(* PLC project Storage_Main, Beckhoff Automation GmbH TwinCAT PLC Control 3.5.13.21 *)
(* stored: creationDateTime 2026-11-24T10:23:53.5609377, modificationDateTime 2026-11-24T10:23:53.5609377 *)

PROGRAM MAIN
// =====================================================================
// MAIN (Structured Text)
// Calls the ST actions and the SFC action ACT_Sequence in a fixed order.
// All variables of the storage system are declared here (HMI uses MAIN.xxx).
// =====================================================================
VAR
    // ---------------- INPUTS ----------------
    B1  AT %I* : BOOL;  // Nr. 5,  B1: reference switch horizontal axis (TRUE = at home)
    B2  AT %I* : BOOL;  // Nr. 6,  B2: light-barrier inside  (TRUE = free, FALSE = pallet)
    B3  AT %I* : BOOL;  // Nr. 7,  B3: light-barrier outside (TRUE = free, FALSE = pallet)
    B4  AT %I* : BOOL;  // Nr. 8,  B4: reference switch vertical axis, top (TRUE = at home)
    B5  AT %I* : BOOL;  // Nr. 11, B5: encoder horizontal axis impulse 1  (EL1202 Term 2 ch. 1)
    B6  AT %I* : BOOL;  // Nr. 12, B6: encoder horizontal axis impulse 2  (EL1202 Term 2 ch. 2)
    B7  AT %I* : BOOL;  // Nr. 13, B7: encoder vertical axis impulse 1    (EL1202 Term 3 ch. 1)
    B8  AT %I* : BOOL;  // Nr. 14, B8: encoder vertical axis impulse 2    (EL1202 Term 3 ch. 2)
    B9  AT %I* : BOOL;  // Nr. 15, B9: reference switch cantilever front (TRUE = arm out)
    B10 AT %I* : BOOL;  // Nr. 16, B10: reference switch cantilever back (TRUE = arm back)

    // ---------------- OUTPUTS ----------------
    M1_Forward AT %Q* : BOOL;  // Nr. 17, Q1 (M1): motor conveyor belt forward
    M1_Back    AT %Q* : BOOL;  // Nr. 18, Q2 (M1): motor conveyor belt backward (moves pallet towards crane)
    M2_Forward AT %Q* : BOOL;  // Nr. 19, Q3 (M2): motor horizontal towards rack
    M2_Back    AT %Q* : BOOL;  // Nr. 20, Q4 (M2): motor horizontal towards conveyor belt
    M3_Down    AT %Q* : BOOL;  // Nr. 21, Q5 (M3): motor vertical axis downward
    M3_Up      AT %Q* : BOOL;  // Nr. 22, Q6 (M3): motor vertical axis upward
    M4_Forward AT %Q* : BOOL;  // Nr. 23, Q7 (M4): motor cantilever forward (arm out)
    M4_Back    AT %Q* : BOOL;  // Nr. 24, Q8 (M4): motor cantilever backward (arm in)

    nTolerance   : DINT := 5;       // Deadband in counts (both axes)

    // ---------------- MANUAL COMMANDS (step S0 only) ----------------
    bJogXForward    : BOOL;         // X towards rack
    bJogXBack       : BOOL;         // X towards conveyor
    bJogYUp         : BOOL;         // Y up
    bJogYDown       : BOOL;         // Y down
    bJogArmOut      : BOOL;         // Arm out (stops at B9)
    bJogArmIn       : BOOL;         // Arm in (stops at B10)
    bJogBeltForward : BOOL;         // Belt moves pallet towards crane (M1_Back, stops when B3 sees a pallet)
    bJogBeltBack    : BOOL;         // Belt moves pallet away from crane (M1_Forward)

    // ---------------- TEACH ----------------
    nTeachSlot : INT := 0;          // 0 = delivery (conveyor), 1..3 = column (X) / row (Y)
    bTeachX    : BOOL;              // Save nPosX into xPosition[nTeachSlot]
    bTeachY    : BOOL;              // Save nPosY into yPosition[nTeachSlot]
    bGoX       : BOOL;              // Move X to xPosition[nTeachSlot]
    bGoY       : BOOL;              // Move Y to yPosition[nTeachSlot]
    nShowX     : DINT;              // Stored X value of nTeachSlot (for HMI)
    nShowY     : DINT;              // Stored Y value of nTeachSlot (for HMI)

    // ---------------- SAVE TAUGHT VALUES (Tc2_Utilities) ----------------
    fbWritePersistent : WritePersistentData;   // Writes all PERSISTENT variables to disk at once
    bSaveData         : BOOL;       // Request: save the persistent data now
    nSaveState        : INT;        // 0 = idle, 1 = start writing, 2 = writing
    bSaveError        : BOOL;       // TRUE if the last write failed
    nLiftOffsetOld    : DINT;       // Last saved nLiftOffset (detects a change from the HMI)
    nLowerOffsetOld   : DINT;       // Last saved nLowerOffset (detects a change from the HMI)

    // ---------------- AUTOMATIC ----------------
    bStartAuto     : BOOL;          // Start automatic mode (homes first)
    bStartHoming   : BOOL;          // Start homing (manual mode)
    bStop          : BOOL;          // Stop everything, back to manual
    bAuto          : BOOL;          // TRUE while automatic mode is active
    bResetSequence : BOOL;          // TRUE for one cycle: ACT_Sequence back to step S0 (STOP / homing timeout)
    SFCReset       : BOOL;          // SFC flag of ACT_Sequence (set from bResetSequence in MAIN)
    nSelColumn     : INT;           // Shelf column to fetch from, chosen by the operator (1..3)
    nSelRow        : INT;           // Shelf row to fetch from, chosen by the operator (1..3)
    bShelfSelected : BOOL;          // Set by the HMI when the operator has chosen a shelf
    bPositionFound : BOOL;          // GRAFCET: PositionFound - target position is loaded (step 71 / 79)
    bInPosition    : BOOL;          // GRAFCET: InPosition - both axes are in position (step 77 / 84)

    // ---------------- POSITIONING ----------------
    nTargetX     : DINT;            // Current X target (GRAFCET: PosX value)
    nTargetY     : DINT;            // Current Y target (GRAFCET: PosY value)
    bDriveX      : BOOL;            // Sequence requests X to move to nTargetX
    bDriveY      : BOOL;            // Sequence requests Y to move to nTargetY
    bPosXReached : BOOL;            // GRAFCET: PosX = TRUE - X has reached nTargetX
    bPosYReached : BOOL;            // GRAFCET: PosY = TRUE - Y has reached nTargetY

    // ---------------- LIMITS ----------------
    nMaxPosX     : DINT := 10000;   // Software end limit X towards rack - MEASURE THIS!
    nMaxPosY     : DINT := 10000;   // Software end limit Y downwards - MEASURE THIS!
    tonHoming    : TON;             // Homing timeout
    bHomingError : BOOL;            // TRUE if a reference switch was not found in time
    tonSettle    : TON;             // 0.5 s settle time at the reference switches

    // ---------------- ENCODER X (B5/B6) ----------------
    nStateX      : BYTE;            // Current state 0..3
    nPrevStateX  : BYTE;            // State in previous cycle
    nPosX        : DINT;            // X position in counts (0 = B1, increases towards rack)
    nErrorCountX : UDINT;           // Number of missed states X

    // ---------------- ENCODER Y (B7/B8) ----------------
    nStateY      : BYTE;            // Current state 0..3
    nPrevStateY  : BYTE;            // State in previous cycle
    nPosY        : DINT;            // Y position in counts (0 = B4 at the top, increases downwards)
    nErrorCountY : UDINT;           // Number of missed states Y

    bInit : BOOL := TRUE;           // First cycle flag (both encoders)

    // ---------------- SEQUENCE / STATUS ----------------
    nStep            : INT := 0;    // Active SFC step number (set by the step actions of ACT_Sequence)
    bHomed           : BOOL;        // TRUE when both axes are homed
    bYTaught         : BOOL;        // TRUE when all Y positions are taught
    bYNotTaught      : BOOL;        // Inverse of bYTaught (for HMI)
    bPalletAtB2      : BOOL;        // TRUE when B2 sees a pallet (HMI lamp)
    bPalletAtB3      : BOOL;        // TRUE when B3 sees a pallet (HMI lamp)
    bShowShelfSelect : BOOL;        // TRUE while the operator must choose a shelf (shows 3x3 on HMI)
    bHideShelfSelect : BOOL;        // Inverse of bShowShelfSelect (hides the 3x3 frame on HMI)
    bSlot0Sel        : BOOL;        // TRUE when teach slot 0 (delivery) is selected (lights the HMI button)
    bSlot1Sel        : BOOL;        // TRUE when teach slot 1 (column 1 / row 1) is selected
    bSlot2Sel        : BOOL;        // TRUE when teach slot 2 (column 2 / row 2) is selected
    bSlot3Sel        : BOOL;        // TRUE when teach slot 3 (column 3 / row 3) is selected
END_VAR

VAR PERSISTENT
    // ---------------- TAUGHT VALUES (kept after power off) ----------------
    // Index 0 = delivery position at the conveyor (GRAFCET: DeliveryPosX / DeliveryPosY)
    // X: [1] = column 1 (nearest conveyor) .. [3] = column 3
    // Y: [1] = row 1 (bottom) .. [3] = row 3 (top). Y counts from the top (B4 = 0) and increases downwards
    xPosition    : ARRAY[0..3] OF DINT := [139, 2995, 5330, 7680];
    yPosition    : ARRAY[0..3] OF DINT := [0, 0, 0, 0];      // MUST BE TAUGHT before automatic mode
    nLiftOffset  : DINT := 30;      // Counts to lift the pallet off the shelf (SFC step S74)
    nLowerOffset : DINT := 50;      // Counts to lower the pallet onto the conveyor (SFC step S86)
END_VAR

            // =====================================================================
// MAIN (Structured Text) - the order of the calls is important:
//   1. ACT_Encoder     (ST)  read the encoders -> nPosX / nPosY
//   2. ACT_Manual      (ST)  status, stop, commands, teach + save, timers,
//                            all motors off, jog in manual mode
//   3. ACT_Sequence    (SFC) homing and the automatic sequence (switches motors ON)
//   4. ACT_Positioning (ST)  drive X / Y to nTargetX / nTargetY
//   5. ACT_Safety      (ST)  end limits and interlocks (always last)
// =====================================================================

ACT_Encoder();
ACT_Manual();

SFCReset := bResetSequence;                 // SFC flag: TRUE = ACT_Sequence back to step S0
ACT_Sequence();                             // SFC: homing and automatic sequence
bResetSequence := FALSE;

// Commands are only accepted in manual mode (step S0). Clear them every cycle,
// so an old button press does not start something later by surprise.
bStartHoming := FALSE;
bStartAuto   := FALSE;
bGoX         := FALSE;
bGoY         := FALSE;

ACT_Positioning();
ACT_Safety();

          

ACTION ACT_Encoder:
                // =====================================================
// ACT_Encoder: count up/down based on the two encoder signals
// X: B5 (A) and B6 (B)    Y: B7 (A) and B8 (B)
// =====================================================
nStateX := 0;                                       // default: A=0, B=0
IF B5 AND NOT B6 THEN nStateX := 1; END_IF          // A=1, B=0
IF B5 AND B6 THEN nStateX := 2; END_IF              // A=1, B=1
IF NOT B5 AND B6 THEN nStateX := 3; END_IF          // A=0, B=1

nStateY := 0;                                       // default: A=0, B=0
IF B7 AND NOT B8 THEN nStateY := 1; END_IF          // A=1, B=0
IF B7 AND B8 THEN nStateY := 2; END_IF              // A=1, B=1
IF NOT B7 AND B8 THEN nStateY := 3; END_IF          // A=0, B=1

IF bInit THEN
    nPrevStateX := nStateX;
    nPrevStateY := nStateY;
    bInit := FALSE;
END_IF

CASE (nStateX + 4 - nPrevStateX) MOD 4 OF
    1: nPosX := nPosX + 1;                          // one step towards rack
    3: nPosX := nPosX - 1;                          // one step towards conveyor
    2: nErrorCountX := nErrorCountX + 1;            // state missed
END_CASE

CASE (nStateY + 4 - nPrevStateY) MOD 4 OF
    1: nPosY := nPosY + 1;                          // one step down
    3: nPosY := nPosY - 1;                          // one step up
    2: nErrorCountY := nErrorCountY + 1;            // state missed
END_CASE

nPrevStateX := nStateX;
nPrevStateY := nStateY;

              
END_ACTION

ACTION ACT_Manual:
                // =====================================================
// ACT_Manual: status, stop, commands, teach + save, timers, jog
// =====================================================

// ---------- 1. STATUS SIGNALS ----------
bPalletAtB2 := NOT B2;                              // light barrier is FALSE when a pallet is in front
bPalletAtB3 := NOT B3;

// Delivery height must be taught, and every shelf row must be low enough to lift nLiftOffset
bYTaught := yPosition[0] > 0 AND yPosition[1] > nLiftOffset AND yPosition[2] > nLiftOffset AND yPosition[3] > nLiftOffset;
bYNotTaught := NOT bYTaught;

bShowShelfSelect := (nStep = 71);
bHideShelfSelect := NOT bShowShelfSelect;
bSlot0Sel := (nTeachSlot = 0);
bSlot1Sel := (nTeachSlot = 1);
bSlot2Sel := (nTeachSlot = 2);
bSlot3Sel := (nTeachSlot = 3);

IF nTeachSlot >= 0 AND nTeachSlot <= 3 THEN
    nShowX := xPosition[nTeachSlot];
    nShowY := yPosition[nTeachSlot];
END_IF


// ---------- 2. STOP: always back to manual mode (step S0) ----------
IF bStop THEN
    bStop := FALSE;
    bStartHoming := FALSE;
    bStartAuto := FALSE;
    bGoX := FALSE;
    bGoY := FALSE;
    bShelfSelected := FALSE;
    bPositionFound := FALSE;
    bInPosition := FALSE;
    bAuto := FALSE;
    bResetSequence := TRUE;                         // ACT_Sequence -> S0 (SFCReset)
END_IF


// ---------- 3. COMMANDS (manual mode only) ----------
// The transitions after step S0 in ACT_Sequence react to the same commands in this cycle.
IF nStep = 0 THEN
    IF bStartHoming THEN
        bHomingError := FALSE;
        bAuto := FALSE;
        bHomed := FALSE;
    END_IF

    IF bStartAuto AND bYTaught THEN                 // Y positions must be taught first
        bHomingError := FALSE;
        bAuto := TRUE;
        bHomed := FALSE;                            // always home before automatic mode
    END_IF

    IF bGoX AND bHomed AND nTeachSlot >= 0 AND nTeachSlot <= 3 THEN
        nTargetX := xPosition[nTeachSlot];
        bPosXReached := FALSE;
    END_IF

    IF bGoY AND bHomed AND nTeachSlot >= 0 AND nTeachSlot <= 3 THEN
        nTargetY := yPosition[nTeachSlot];
        bPosYReached := FALSE;
    END_IF
END_IF


// ---------- 4. TEACH: save current position into the arrays (manual mode only) ----------
IF bTeachX THEN
    bTeachX := FALSE;
    IF nStep = 0 AND bHomed AND nTeachSlot >= 0 AND nTeachSlot <= 3 THEN
        xPosition[nTeachSlot] := nPosX;
        bSaveData := TRUE;                          // write to disk at once
    END_IF
END_IF

IF bTeachY THEN
    bTeachY := FALSE;
    IF nStep = 0 AND bHomed AND nTeachSlot >= 0 AND nTeachSlot <= 3 THEN
        yPosition[nTeachSlot] := nPosY;
        bSaveData := TRUE;                          // write to disk at once
    END_IF
END_IF

// Lift / lower offset changed on the HMI -> save as well
IF nLiftOffset <> nLiftOffsetOld OR nLowerOffset <> nLowerOffsetOld THEN
    nLiftOffsetOld := nLiftOffset;
    nLowerOffsetOld := nLowerOffset;
    bSaveData := TRUE;
END_IF


// ---------- 5. SAVE: write the PERSISTENT variables to disk (survives a power cut) ----------
// WritePersistentData starts on a rising edge of START. nSaveState makes sure that
// START is TRUE until the write has started, and FALSE again before the next write.
CASE nSaveState OF
    0:  // idle: wait for a save request
        IF bSaveData THEN
            bSaveData := FALSE;
            nSaveState := 1;
        END_IF

    1:  // START = TRUE: wait until the write has started (or failed at once)
        IF fbWritePersistent.BUSY OR fbWritePersistent.ERR THEN
            nSaveState := 2;
        END_IF

    2:  // START = FALSE: wait until the write is finished
        IF NOT fbWritePersistent.BUSY THEN
            nSaveState := 0;
        END_IF
END_CASE

fbWritePersistent(NETID := '', PORT := 851, START := (nSaveState = 1), TMOUT := T#5S, MODE := SPDM_2PASS);
bSaveError := fbWritePersistent.ERR;


// ---------- 6. TIMERS (called every cycle so they reset themselves) ----------
tonHoming(IN := (nStep = 10 OR nStep = 11), PT := T#20S);
tonSettle(IN := (nStep = 12), PT := T#500MS);

IF tonHoming.Q THEN
    bHomingError := TRUE;
    bAuto := FALSE;
    bResetSequence := TRUE;                         // ACT_Sequence -> S0, motors off
END_IF


// ---------- 7. MOTORS OFF + JOG ----------
// Default: all motors off. ACT_Sequence (called after this action) switches on what
// the active step needs. In manual mode (S0) the jog buttons are used.
M1_Forward := FALSE;
M1_Back    := FALSE;
M2_Forward := FALSE;
M2_Back    := FALSE;
M3_Down    := FALSE;
M3_Up      := FALSE;
M4_Forward := FALSE;
M4_Back    := FALSE;
bDriveX    := FALSE;
bDriveY    := FALSE;

IF nStep = 0 THEN
    M2_Forward := bJogXForward AND NOT bJogXBack;
    M2_Back    := bJogXBack AND NOT bJogXForward;
    M3_Down    := bJogYDown AND NOT bJogYUp;
    M3_Up      := bJogYUp AND NOT bJogYDown;
    M4_Forward := bJogArmOut AND NOT bJogArmIn;
    M4_Back    := bJogArmIn AND NOT bJogArmOut;
    M1_Back    := bJogBeltForward AND NOT bJogBeltBack AND B3;   // stops when B3 sees a pallet
    M1_Forward := bJogBeltBack AND NOT bJogBeltForward;
END_IF

              
END_ACTION

ACTION ACT_Positioning:
                // =====================================================
// ACT_Positioning: drive X and Y to their targets
// =====================================================
// An axis stops for good when it is within the tolerance (bPosXReached / bPosYReached),
// so it does not hunt back and forth if the motor coasts a little.
IF bDriveX AND NOT bPosXReached THEN
    IF nPosX < nTargetX - nTolerance THEN
        M2_Forward := TRUE;                         // towards rack
    END_IF
    IF nPosX > nTargetX + nTolerance THEN
        M2_Back := TRUE;                            // towards conveyor
    END_IF
    IF NOT M2_Forward AND NOT M2_Back THEN
        bPosXReached := TRUE;
    END_IF
END_IF

IF bDriveY AND NOT bPosYReached THEN
    IF nPosY < nTargetY - nTolerance THEN
        M3_Down := TRUE;                            // larger Y = further down
    END_IF
    IF nPosY > nTargetY + nTolerance THEN
        M3_Up := TRUE;                              // smaller Y = further up
    END_IF
    IF NOT M3_Down AND NOT M3_Up THEN
        bPosYReached := TRUE;
    END_IF
END_IF

              
END_ACTION

ACTION ACT_Safety:
                // =====================================================
// ACT_Safety: end limits and interlocks (always called last)
// =====================================================
// X: hardware end at the conveyor (B1)
IF B1 THEN
    M2_Back := FALSE;
END_IF

// X: software end towards the rack
IF bHomed AND nPosX >= nMaxPosX THEN
    M2_Forward := FALSE;
END_IF

// X may only move when the arm is back (B10)
IF NOT B10 THEN
    M2_Forward := FALSE;
    M2_Back    := FALSE;
END_IF

// Y: hardware end at the top (B4)
IF B4 THEN
    M3_Up := FALSE;
END_IF

// Y: software end at the bottom
IF bHomed AND nPosY >= nMaxPosY THEN
    M3_Down := FALSE;
END_IF

// Arm: end positions
IF B9 THEN
    M4_Forward := FALSE;
END_IF

IF B10 THEN
    M4_Back := FALSE;
END_IF

// Never both directions at the same time
IF M1_Forward AND M1_Back THEN
    M1_Forward := FALSE;
    M1_Back    := FALSE;
END_IF

IF M2_Forward AND M2_Back THEN
    M2_Forward := FALSE;
    M2_Back    := FALSE;
END_IF

IF M3_Down AND M3_Up THEN
    M3_Down := FALSE;
    M3_Up   := FALSE;
END_IF

IF M4_Forward AND M4_Back THEN
    M4_Forward := FALSE;
    M4_Back    := FALSE;
END_IF

              
END_ACTION

ACTION ACT_Sequence:
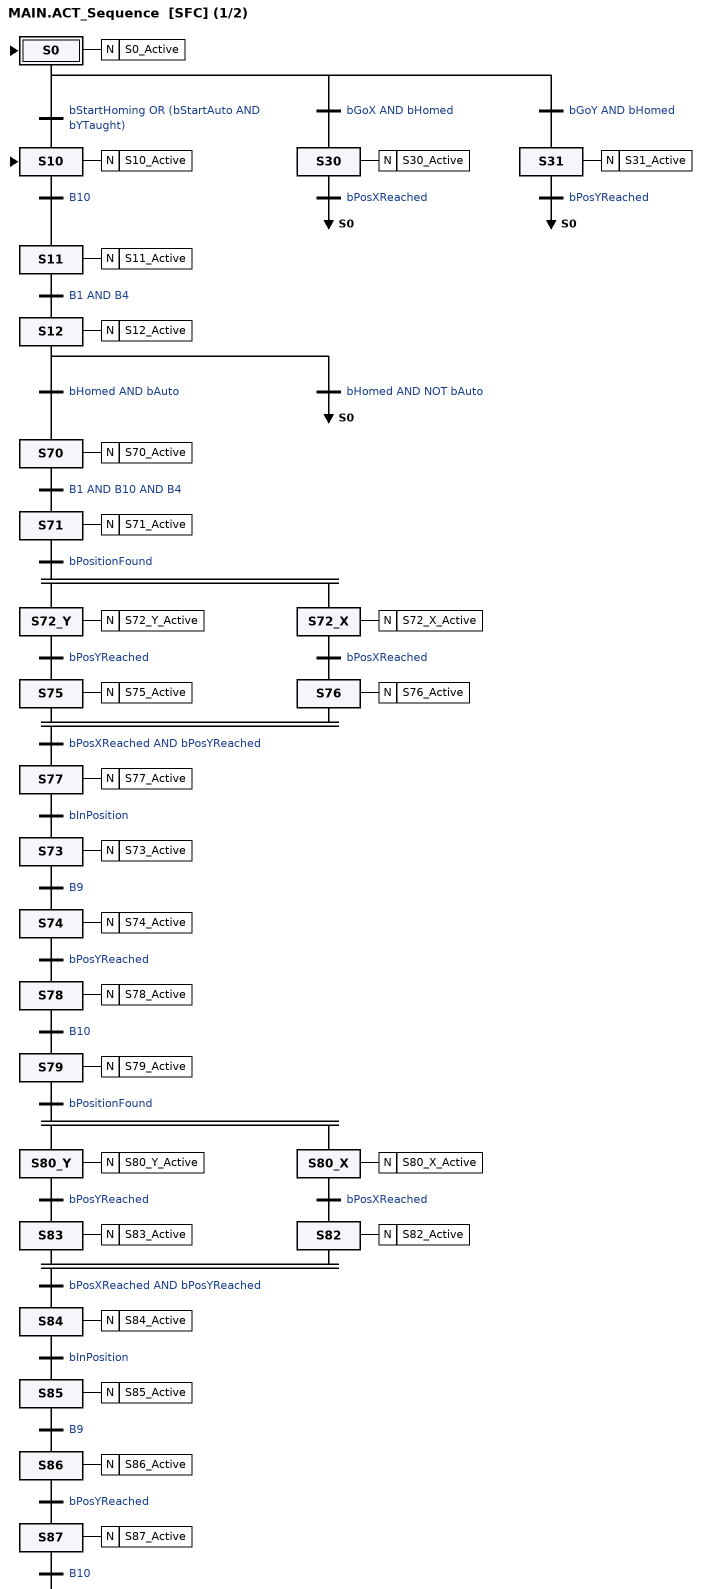
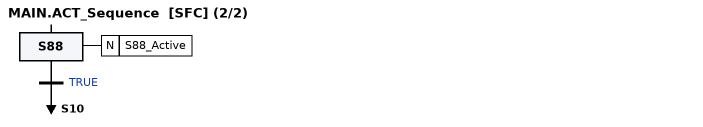
INITIAL_STEP S0:
  S0_Active(N);
END_STEP
TRANSITION FROM S0 TO S10
  := bStartHoming OR (bStartAuto AND bYTaught);
END_TRANSITION
TRANSITION FROM S0 TO S30
  := bGoX AND bHomed;
END_TRANSITION
TRANSITION FROM S0 TO S31
  := bGoY AND bHomed;
END_TRANSITION
STEP S10:
  S10_Active(N);
END_STEP
TRANSITION FROM S10 TO S11
  := B10;
END_TRANSITION
STEP S11:
  S11_Active(N);
END_STEP
TRANSITION FROM S11 TO S12
  := B1 AND B4;
END_TRANSITION
STEP S12:
  S12_Active(N);
END_STEP
TRANSITION FROM S12 TO S70
  := bHomed AND bAuto;
END_TRANSITION
TRANSITION FROM S12 TO S0
  := bHomed AND NOT bAuto;
END_TRANSITION
STEP S70:
  S70_Active(N);
END_STEP
TRANSITION FROM S70 TO S71
  := B1 AND B10 AND B4;
END_TRANSITION
STEP S71:
  S71_Active(N);
END_STEP
TRANSITION FROM S71 TO (S72_Y, S72_X)
  := bPositionFound;
END_TRANSITION
STEP S72_Y:
  S72_Y_Active(N);
END_STEP
TRANSITION FROM S72_Y TO S75
  := bPosYReached;
END_TRANSITION
STEP S75:
  S75_Active(N);
END_STEP
TRANSITION FROM (S75, S76) TO S77
  := bPosXReached AND bPosYReached;
END_TRANSITION
STEP S72_X:
  S72_X_Active(N);
END_STEP
TRANSITION FROM S72_X TO S76
  := bPosXReached;
END_TRANSITION
STEP S76:
  S76_Active(N);
END_STEP
STEP S77:
  S77_Active(N);
END_STEP
TRANSITION FROM S77 TO S73
  := bInPosition;
END_TRANSITION
STEP S73:
  S73_Active(N);
END_STEP
TRANSITION FROM S73 TO S74
  := B9;
END_TRANSITION
STEP S74:
  S74_Active(N);
END_STEP
TRANSITION FROM S74 TO S78
  := bPosYReached;
END_TRANSITION
STEP S78:
  S78_Active(N);
END_STEP
TRANSITION FROM S78 TO S79
  := B10;
END_TRANSITION
STEP S79:
  S79_Active(N);
END_STEP
TRANSITION FROM S79 TO (S80_Y, S80_X)
  := bPositionFound;
END_TRANSITION
STEP S80_Y:
  S80_Y_Active(N);
END_STEP
TRANSITION FROM S80_Y TO S83
  := bPosYReached;
END_TRANSITION
STEP S83:
  S83_Active(N);
END_STEP
TRANSITION FROM (S83, S82) TO S84
  := bPosXReached AND bPosYReached;
END_TRANSITION
STEP S80_X:
  S80_X_Active(N);
END_STEP
TRANSITION FROM S80_X TO S82
  := bPosXReached;
END_TRANSITION
STEP S82:
  S82_Active(N);
END_STEP
STEP S84:
  S84_Active(N);
END_STEP
TRANSITION FROM S84 TO S85
  := bInPosition;
END_TRANSITION
STEP S85:
  S85_Active(N);
END_STEP
TRANSITION FROM S85 TO S86
  := B9;
END_TRANSITION
STEP S86:
  S86_Active(N);
END_STEP
TRANSITION FROM S86 TO S87
  := bPosYReached;
END_TRANSITION
STEP S87:
  S87_Active(N);
END_STEP
TRANSITION FROM S87 TO S88
  := B10;
END_TRANSITION
STEP S88:
  S88_Active(N);
END_STEP
TRANSITION FROM S88 TO S10
  := TRUE;
END_TRANSITION
STEP S30:
  S30_Active(N);
END_STEP
TRANSITION FROM S30 TO S0
  := bPosXReached;
END_TRANSITION
STEP S31:
  S31_Active(N);
END_STEP
TRANSITION FROM S31 TO S0
  := bPosYReached;
END_TRANSITION
END_ACTION

ACTION S0_Active:
                // S0: Manual mode (initial step)
// Jog, teach and the commands are handled in MAIN (ST) while nStep = 0.
nStep := 0;
              
END_ACTION

ACTION S10_Active:
                // S10: Homing - arm back (until B10)
nStep := 10;
bHomed := FALSE;
M4_Back := TRUE;
              
END_ACTION

ACTION S11_Active:
                // S11: Homing - X to B1 and Y to B4 at the same time
nStep := 11;
M2_Back := NOT B1;                     // each axis stops at its own switch
M3_Up   := NOT B4;
              
END_ACTION

ACTION S12_Active:
                // S12: Homing - wait 0.5 s (tonSettle in MAIN), then set both positions to 0
nStep := 12;
IF tonSettle.Q THEN
    nPosX := 0;
    nPosY := 0;
    bHomed := TRUE;
END_IF
              
END_ACTION

ACTION S70_Active:
                // S70 = E70 Entry step: wait until the crane is at home (B1 * B10 * B4)
nStep := 70;
bShelfSelected := FALSE;                    // ignore any old shelf selection
              
END_ACTION

ACTION S71_Active:
                // S71: Get PosX and PosY from the arrays according to the operator's choice
// (nStep = 71 shows the 3x3 shelf selection on the HMI)
nStep := 71;
bPosXReached := FALSE;
bPosYReached := FALSE;

IF bShelfSelected THEN
    bShelfSelected := FALSE;
    IF nSelColumn >= 1 AND nSelColumn <= 3 AND nSelRow >= 1 AND nSelRow <= 3 THEN
        nTargetX := xPosition[nSelColumn];
        nTargetY := yPosition[nSelRow];
        bPositionFound := TRUE;
    END_IF
END_IF
              
END_ACTION

ACTION S72_Y_Active:
                // S72 (Y part): Y moves to the shelf height (M3_Down via ACT_Positioning)
nStep := 72;
bPositionFound := FALSE;
bDriveY := TRUE;
              
END_ACTION

ACTION S75_Active:
                // S75: Y in position (M3 off), waits for X
nStep := 75;
              
END_ACTION

ACTION S72_X_Active:
                // S72 (X part): X moves to the shelf column (M2_Forward via ACT_Positioning)
nStep := 72;
bPositionFound := FALSE;
bDriveX := TRUE;
              
END_ACTION

ACTION S76_Active:
                // S76: X in position (M2 off), waits for Y
nStep := 76;
              
END_ACTION

ACTION S77_Active:
                // S77: Both axes in position
nStep := 77;
bInPosition := TRUE;
              
END_ACTION

ACTION S73_Active:
                // S73: Arm out under the pallet (until B9)
nStep := 73;
M4_Forward := TRUE;
bInPosition := FALSE;
nTargetY := yPosition[nSelRow] - nLiftOffset;   // prepare the lift (up = smaller Y)
bPosYReached := FALSE;
              
END_ACTION

ACTION S74_Active:
                // S74: Lift the pallet off the shelf (M3_Up via ACT_Positioning)
nStep := 74;
bDriveY := TRUE;
              
END_ACTION

ACTION S78_Active:
                // S78: Arm back with the pallet (until B10)
nStep := 78;
M4_Back := TRUE;
              
END_ACTION

ACTION S79_Active:
                // S79: Get the delivery position (index 0 = conveyor)
nStep := 79;
nTargetX := xPosition[0];              // DeliveryPosX
nTargetY := yPosition[0];              // DeliveryPosY
bPosXReached := FALSE;
bPosYReached := FALSE;
bPositionFound := TRUE;
              
END_ACTION

ACTION S80_Y_Active:
                // S80/S81 (Y part): Y moves up or down to the delivery height.
// ACT_Positioning chooses the direction (M3_Up or M3_Down) by itself.
nStep := 80;
bPositionFound := FALSE;
bDriveY := TRUE;
              
END_ACTION

ACTION S83_Active:
                // S83: Y in position (M3 off), waits for X
nStep := 83;
              
END_ACTION

ACTION S80_X_Active:
                // S80/S81 (X part): X moves back to the conveyor (M2_Back via ACT_Positioning)
nStep := 80;
bPositionFound := FALSE;
bDriveX := TRUE;
              
END_ACTION

ACTION S82_Active:
                // S82: X in position (M2 off), waits for Y
nStep := 82;
              
END_ACTION

ACTION S84_Active:
                // S84: Both axes in position
nStep := 84;
bInPosition := TRUE;
              
END_ACTION

ACTION S85_Active:
                // S85: Arm out over the conveyor (until B9)
nStep := 85;
M4_Forward := TRUE;
bInPosition := FALSE;
nTargetY := yPosition[0] + nLowerOffset;   // prepare lowering (down = larger Y)
bPosYReached := FALSE;
              
END_ACTION

ACTION S86_Active:
                // S86: Lower the pallet onto the conveyor (M3_Down via ACT_Positioning)
nStep := 86;
bDriveY := TRUE;
              
END_ACTION

ACTION S87_Active:
                // S87: Arm back (until B10)
nStep := 87;
M4_Back := TRUE;
              
END_ACTION

ACTION S88_Active:
                // S88 = S70 Exit step: home again. Homing returns to S70 because bAuto is still TRUE.
nStep := 88;
              
END_ACTION

ACTION S30_Active:
                // S30: Manual - move X to xPosition[nTeachSlot] (target set in ACT_Manual)
nStep := 30;
bDriveX := TRUE;
              
END_ACTION

ACTION S31_Active:
                // S31: Manual - move Y to yPosition[nTeachSlot] (target set in ACT_Manual)
nStep := 31;
bDriveY := TRUE;
              
END_ACTION
END_PROGRAM
